// TIA Portal V21 export
VAR_GLOBAL   // PLC tag table "IO_horizontale Achse"
   ModePos_h AT %MW1 : Int;   //    {ExternalAccessible false}
   AxisEnabled_h AT %M3.4 : Bool;
   AxisPosOK_h AT %M3.0 : Bool;
   AxisRef_h AT %M3.1 : Bool;
   AxisError_h AT %M3.2 : Bool;
   Error_h AT %M3.3 : Bool;
   ActVel_h AT %M23.0 : LReal;
   ActPos_h AT %M32.0 : LReal;
END_VAR
